{attribute 'qualified_only'}
{attribute 'strict'}
TYPE E_Recipe_Root_Folder :
(
	PLC := 0,
	Develop_1,
	Develop_2,
	Develop_3,
	Develop_4	
);
END_TYPE

(* stored: Version 1.1.0.1, ProductVersion 3.1.4024.12
   DUT E_Recipe_Root_Folder: Id {951518db-2f03-4c7a-a91a-5816ff396c59} *)
